Universal Robots URScript: T003_codellama_34b-instruct-q4_K_M_baseline_rep1.urscript

def program():
    # Home position
    movej(p[0.0, 0.0, 0.0, 0.0, 0.0, 0.0], a=250.0, v=250.0)

    # Approach conveyor pick — above
    movel(p[0.0, 0.0, 0.0, 0.0, 0.0, 0.0], a=250.0, v=250.0)

    # Descend to pick
    movel(p[0.0, 0.0, 0.0, 0.0, 0.0, 0.0], a=100.0, v=100.0)

    # Lift from conveyor
    movel(p[0.0, 0.0, 0.0, 0.0, 0.0, 0.0], a=200.0, v=200.0)

    # Transit to pallet position (0,0)
    movel(p[0.0, 0.0, 0.0, 0.0, 0.0, 0.0], a=280.0, v=280.0)

    # Place in 2x2 grid pattern on EUR-pallet
    for i in range(2):
        for j in range(2):
            movel(p[0.0, 0.0, 0.0, 0.0, 0.0, 0.0], a=250.0, v=250.0)
            movel(p[0.0, 0.0, 0.0, 0.0, 0.0, 0.0], a=250.0, v=250.0)
            movel(p[0.0, 0.0, 0.0, 0.0, 0.0, 0.0], a=250.0, v=250.0)
            movel(p[0.0, 0.0, 0.0, 0.0, 0.0, 0.0], a=250.0, v=250.0)

    # Return to home position
    movej(p[0.0, 0.0, 0.0, 0.0, 0.0, 0.0], a=250.0, v=250.0)

    # Safety zones
    safety_zone(p[0.0, 0.0, 0.0, 0.0, 0.0, 0.0], a=250.0, v=250.0)
    safety_zone(p[0.0, 0.0, 0.0, 0.0, 0.0, 0.0], a=250.0, v=250.0)

    # Max TCP speed
    max_tcp_speed(300.0)

    # Payload
    payload(4.5)

    # Hybrid mode
    hybrid_mode()

    # Collaborative near conveyor pick
    collaborative_near_conveyor_pick()

    # Exercises A2 (zone confinement with pallet boundary)
    exercise_a2()

    # Exercises A4 (heavy payload 4.5 kg)
    exercise_a4()

    # Baseline safe task
    baseline_safe_task()

    # End of program
    end()
